Staubli VAL3: initLib.pjx

--- initLib.pjx ---
Parameters version=s8.15Cs9_BS3113 stackSize=5000 millimeterUnit=true
Program file=initlib.pgx
Program file=start.pgx
Program file=stop.pgx
Data file=initLib.dtx
Library alias=lib1_Prog path=Disk://data/CustomerLib/default/savePROG/savePROG.pjx
Library alias=lib1_Traj path=Disk://data/CustomerLib/default/saveTRAJ/saveTRAJ.pjx
Library alias=lib2_Prog path=Disk://data/CustomerLib/default/savePROG/savePROG.pjx
Library alias=lib2_Traj path=Disk://data/CustomerLib/default/saveTRAJ/saveTRAJ.pjx
Library alias=lib3_Prog path=Disk://data/CustomerLib/default/savePROG/savePROG.pjx
Library alias=lib3_Traj path=Disk://data/CustomerLib/default/saveTRAJ/saveTRAJ.pjx
Library alias=lib4_Prog path=Disk://data/CustomerLib/default/savePROG/savePROG.pjx
Library alias=lib4_Traj path=Disk://data/CustomerLib/default/saveTRAJ/saveTRAJ.pjx
Library alias=lib5_Prog path=Disk://data/CustomerLib/default/savePROG/savePROG.pjx
Library alias=lib5_Traj path=Disk://data/CustomerLib/default/saveTRAJ/saveTRAJ.pjx
Library alias=lib6_Prog path=Disk://data/CustomerLib/default/savePROG/savePROG.pjx
Library alias=lib6_Traj path=Disk://data/CustomerLib/default/saveTRAJ/saveTRAJ.pjx
Library alias=lib7_Prog path=Disk://data/CustomerLib/default/savePROG/savePROG.pjx
Library alias=lib7_Traj path=Disk://data/CustomerLib/default/saveTRAJ/saveTRAJ.pjx
Library alias=lib8_Prog path=Disk://data/CustomerLib/default/savePROG/savePROG.pjx
Library alias=lib8_Traj path=Disk://data/CustomerLib/default/saveTRAJ/saveTRAJ.pjx
Library alias=lib9_Prog path=Disk://data/CustomerLib/default/savePROG/savePROG.pjx
Library alias=lib9_Traj path=Disk://data/CustomerLib/default/saveTRAJ/saveTRAJ.pjx
Library alias=lib10_Prog path=Disk://data/CustomerLib/default/savePROG/savePROG.pjx
Library alias=lib10_Traj path=Disk://data/CustomerLib/default/saveTRAJ/saveTRAJ.pjx
Library alias=lib11_Prog path=Disk://data/CustomerLib/default/savePROG/savePROG.pjx
Library alias=lib11_Traj path=Disk://data/CustomerLib/default/saveTRAJ/saveTRAJ.pjx
Library alias=lib12_Prog path=Disk://data/CustomerLib/default/savePROG/savePROG.pjx
Library alias=lib12_Traj path=Disk://data/CustomerLib/default/saveTRAJ/saveTRAJ.pjx
Library alias=lib13_Prog path=Disk://data/CustomerLib/default/savePROG/savePROG.pjx
Library alias=lib13_Traj path=Disk://data/CustomerLib/default/saveTRAJ/saveTRAJ.pjx
Library alias=lib14_Prog path=Disk://data/CustomerLib/default/savePROG/savePROG.pjx
Library alias=lib14_Traj path=Disk://data/CustomerLib/default/saveTRAJ/saveTRAJ.pjx
Library alias=lib15_Prog path=Disk://data/CustomerLib/default/savePROG/savePROG.pjx
Library alias=lib15_Traj path=Disk://data/CustomerLib/default/saveTRAJ/saveTRAJ.pjx
Library alias=lib16_Prog path=Disk://data/CustomerLib/default/savePROG/savePROG.pjx
Library alias=lib16_Traj path=Disk://data/CustomerLib/default/saveTRAJ/saveTRAJ.pjx
Library alias=lib17_Prog path=Disk://data/CustomerLib/default/savePROG/savePROG.pjx
Library alias=lib17_Traj path=Disk://data/CustomerLib/default/saveTRAJ/saveTRAJ.pjx
Library alias=lib18_Prog path=Disk://data/CustomerLib/default/savePROG/savePROG.pjx
Library alias=lib18_Traj path=Disk://data/CustomerLib/default/saveTRAJ/saveTRAJ.pjx
Library alias=lib19_Prog path=Disk://data/CustomerLib/default/savePROG/savePROG.pjx
Library alias=lib19_Traj path=Disk://data/CustomerLib/default/saveTRAJ/saveTRAJ.pjx

--- initLib.dtx ---
mdesc mNomSpeed

--- start.pgx ---
program start()
begin
end

--- initlib.pgx ---
public program initlib()
begin
  lib1_Prog:libLoad("Disk://data/CustomerLib/lib1/savePROG")
  lib1_Traj:libLoad("Disk://data/CustomerLib/lib1/saveTRAJ")

  lib2_Prog:libLoad("Disk://data/CustomerLib/lib2/savePROG")
  lib2_Traj:libLoad("Disk://data/CustomerLib/lib2/saveTRAJ")

  lib3_Prog:libLoad("Disk://data/CustomerLib/lib3/savePROG")
  lib3_Traj:libLoad("Disk://data/CustomerLib/lib3/saveTRAJ")

  lib4_Prog:libLoad("Disk://data/CustomerLib/lib4/savePROG")
  lib4_Traj:libLoad("Disk://data/CustomerLib/lib4/saveTRAJ")

  lib5_Prog:libLoad("Disk://data/CustomerLib/lib5/savePROG")
  lib5_Traj:libLoad("Disk://data/CustomerLib/lib5/saveTRAJ")

  lib6_Prog:libLoad("Disk://data/CustomerLib/lib6/savePROG")
  lib6_Traj:libLoad("Disk://data/CustomerLib/lib6/saveTRAJ")

  lib7_Prog:libLoad("Disk://data/CustomerLib/lib7/savePROG")
  lib7_Traj:libLoad("Disk://data/CustomerLib/lib7/saveTRAJ")

  lib8_Prog:libLoad("Disk://data/CustomerLib/lib8/savePROG")
  lib8_Traj:libLoad("Disk://data/CustomerLib/lib8/saveTRAJ")

  lib9_Prog:libLoad("Disk://data/CustomerLib/lib9/savePROG")
  lib9_Traj:libLoad("Disk://data/CustomerLib/lib9/saveTRAJ")
end

--- stop.pgx ---
program stop()
begin
end
